KUKA KRL program: Feature.src

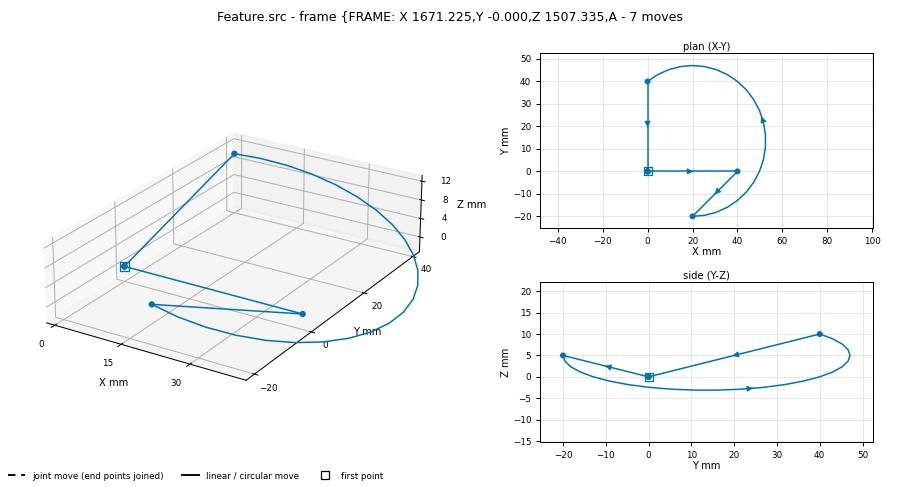
[picture p0: tool path of Feature.src in frame {FRAME: X 1671.225,Y -0.000,Z 1507.335,A, 7 of 13 moves have a stored position in this frame; points joined in program order, loops and branches not executed]
DEF Feature()
; Program generated by RoboDK v5.9.4 for R1 on 26/10/2026 01:01:11
; Using nominal kinematics.
BAS(#INITMOV,0)
$ORI_TYPE  = #VAR
$CIRC_TYPE = #BASE
$VEL.ORI1 = 200
$VEL.ORI2 = 200
$ACC.ORI1 = 100
$ACC.ORI2 = 100
$ADVANCE = 2
$ACT_EX_AX = 0
PTP $AXIS_ACT ; skip BCO quickly
$BASE = {FRAME: X 1671.225,Y -0.000,Z 1507.335,A 30.000,B 0.000,C 0.000}
$TOOL = {FRAME: X 0.000,Y 0.000,Z 120.000,A 0.000,B 15.000,C 0.000}
;------ Using Tool frame number 1 ------
$ACT_TOOL = 1
$TOOL=TOOL_DATA[1]
;------ $TOOL = {FRAME: X 0.000,Y 0.000,Z 120.000,A 0.000,B 15.000,C 0.000}
PTP {AXIS: A1 -0.000,A2 -90.000,A3 100.000,A4 0.000,A5 35.000,A6 90.000}
; PTP {POS:X 1586.372,Y 0.000,Z 1592.188,A -90.000,B -0.000,C -135.000,S 'B010',T 'B000011'}
$VEL.CP = 0.25000
$APO.CPTP = 5
$APO.CDIS = 5
PTP {POS:X 0.000,Y 0.000,Z 0.000,A -130.729,B -10.545,C -134.007} C_PTP
LIN {X 40.000,Y 0.000,Z 0.000,A -130.729,B -10.545,C -134.007} C_DIS
LIN {X 20.000,Y -20.000,Z 5.000,A -130.729,B -10.545,C -134.007} C_DIS
CIRC {X 40.000,Y 40.000,Z 0.000},{X 0.000,Y 40.000,Z 10.000,A -130.729,B -10.545,C -134.007} C_DIS
$ACC.CP = 0.800
$VEL.CP = 0.12000
LIN {X 0.000,Y 0.000,Z 0.000,A -130.729,B -10.545,C -134.007}
LIN {X 0.000,Y 0.000,Z 0.000,A -144.509,B 4.006,C -133.211}
PTP {POS:X 0.000,Y 0.000,Z 0.000,A -130.729,B -10.545,C -134.007}
$ACC.CP = 1.500
$VEL.CP = 0.30000
$ACC.CP = 0.050
$OUT[5] = TRUE
$OUT[3] = FALSE
WAIT FOR $IN[2]==TRUE
; use custom post processor to support timeout
WAIT FOR $IN[4]==FALSE
WAIT SEC 1.500
HALT
; A comment line
Wait for StrClear($LOOP_MSG[])
$LOOP_CONT = TRUE
$LOOP_MSG[] = "A message"
WAIT FOR NOT $LOOP_CONT
SubProg()
SpacedName()
ExternalProg()
Long_ProgramName12()
AnotherLong_ExternalName()
SetRPM700
Ab_c()
custom_code(1)
ThreadProg()
$OUT[2] = 3.5
;------ Using Reference frame number 2 ------
$ACT_BASE = 2
$BASE=BASE_DATA[2]
;------ $BASE = {FRAME: X 1711.225,Y -30.000,Z 1527.335,A 0.000,B 0.000,C 0.000}
$TOOL = {FRAME: X 10.000,Y 0.000,Z 150.000,A 0.000,B 0.000,C 0.000}
PTP {POS:X -40.000,Y 30.000,Z -40.000,A -100.729,B -10.545,C -134.007}
PTP {AXIS: A1 -0.000,A2 -90.000,A3 100.000,A4 0.000,A5 35.000,A6 90.000}
; PTP {POS:X 1586.372,Y 0.000,Z 1592.188,A -90.000,B -0.000,C -135.000,S 'B010',T 'B000011'}
LIN {X -53.660,Y 35.176,Z -26.340,A -100.729,B -10.545,C -134.007}
;------ Using Tool frame number 1 ------
$ACT_TOOL = 1
$TOOL=TOOL_DATA[1]
;------ $TOOL = {FRAME: X 0.000,Y 0.000,Z 120.000,A 0.000,B 15.000,C 0.000}
$BASE = {FRAME: X 1671.225,Y -0.000,Z 1507.335,A 30.000,B 0.000,C 0.000}
PTP {AXIS: A1 -0.000,A2 -90.000,A3 100.000,A4 0.000,A5 35.000,A6 90.000}
; PTP {POS:X 1586.372,Y 0.000,Z 1592.188,A -90.000,B -0.000,C -135.000,S 'B010',T 'B000011'}
END
